// TIA Portal V21 export
FUNCTION_BLOCK "LockedSafety"   // FB1, F_FBD
{ S7_Optimized_Access := 'TRUE' }
// Main safety block of a safety program with a password.
   VAR
      source : Bool;
      target : Bool;
   END_VAR
BEGIN

REGION Network 1: Copy
   // Copies one bit to another.
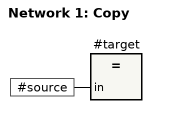
   #target := #source;
END_REGION
END_FUNCTION_BLOCK
